{attribute 'no_assign'}
FUNCTION_BLOCK FB_DO_WTURBINE_LD0_WPPD1_DevOp EXTENDS FB_AcsiCommonDataClass
VAR_INPUT
	st_: FB_DO_WTURBINE_LD0_WPPD1_DevOp_st := (sObjectName:='st', sClass:='ENC', bLinkResult:=THIS^.AddDataToContainer(ipData:=st_));
END_VAR
VAR
END_VAR

END_FUNCTION_BLOCK

(* stored: Version 1.1.0.1
   POU FB_DO_WTURBINE_LD0_WPPD1_DevOp: Id {0f22ed42-39d7-437f-b548-927c5b4bf6b1}, SpecialFunc None *)
